// TIA Portal V21 export
// export: Created 2026-11-11T00:47:15.7506712Z, ExportSetting WithDefaults, DisplayName Totally Integrated Automation Portal, DisplayVersion V21 Update 3, DisplayName STEP 7 Professional, DisplayVersion V21 Update 3, DisplayName STEP 7 Safety, DisplayVersion V21, DisplayName Tech WebApplication, DisplayVersion V21, DisplayName WinCC Basic/Comfort/Advanced, DisplayVersion V21 Update 3, DisplayName WinCC Unified, DisplayVersion V21 Update 3
FUNCTION_BLOCK "FB_Fbd_ex040"   // FB83, FBD
{ S7_Optimized_Access := 'TRUE' }
VERSION : 0.1
// stored: AutoNumber true, IsIECCheckEnabled false, IsRetainMemResEnabled false, MemoryReserve 100, SetENOAutomatically false, UDAEnableTagReadback false
   VAR_INPUT
      v_size : DInt;
   END_VAR
   VAR_OUTPUT
      v_ret_val : WString;
   END_VAR
BEGIN

REGION Network 1: GetBlockName - Read out name of the block
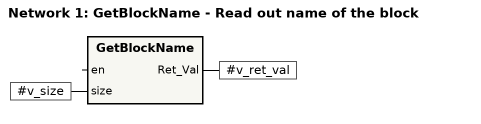
   #v_ret_val := GetBlockName(size := #v_size);
END_REGION
END_FUNCTION_BLOCK
